// Float field value of a typed publisher (PublishLREAL), BROTLib#4: LREAL_TO_STRING with no 'i', so a whole number
// (15.0 prints '15') stays a float. Empty for NaN and infinity: line protocol has no such value, the caller does not
// publish the point.
FUNCTION F_InfluxFloatValue : STRING(255)
VAR_INPUT
	fValue		: LREAL;
END_VAR
VAR
	nBits		: ULINT;
END_VAR

// NaN and infinity have all exponent bits set. Read the bits instead of comparing: a comparison with NaN is an invalid
// floating point operation, which stops the PLC (TcUnit never reported completion in CI).
MEMCPY(ADR(nBits), ADR(fValue), SIZEOF(nBits));
IF (nBits AND 16#7FF0000000000000) = 16#7FF0000000000000 THEN
	F_InfluxFloatValue := '';
ELSE
	F_InfluxFloatValue := LREAL_TO_STRING(fValue);
END_IF

END_FUNCTION

(* stored: Version 1.1.0.1, ProductVersion 3.1.4024.15
   POU F_InfluxFloatValue: Id {65e837f0-c051-429a-90a9-2430d071b0b9}, SpecialFunc None *)
